(* Tests the contract between a caller's batch and a log exporter. *)
FUNCTION_BLOCK FB_TestLogExporters EXTENDS FB_TestSuite

THIS^.testExportSerializesWholeBatch();

(*
	export takes ownership of every record in the caller's batch and passes them to the serializer, so the
	caller holds nothing the exporter will release. Grouping by resource and scope is tested in FB_TestProtoJsonSerializer.
*)
METHOD testExportSerializesWholeBatch : REFERENCE TO FB_Test
VAR CONSTANT
	RECORD_COUNT: UDINT := 2;  // more than one, so the whole batch has to move, not just its head
END_VAR
VAR
	resource: FB_Resource(schemaUrl:='');
	provider: FB_LoggerProvider(resource:=resource);
	scope: FB_InstrumentationScope(name:='exporter.test', version:='1.0.0', schemaUrl:='');
	logger: FB_Logger(scope:=scope, provider:=provider);
	processor: FB_LogRecordProcessor_ForRecordsInspection(
		maxQueueSize:=0,
		scheduledDelayMillis:=1000,
		maxExportBatchSize:=512,
		exporter:=0
	);
	exporter: FB_LogRecordExporter_File_ForSerializationInspection;
	serialized: REFERENCE TO FB_LogRecordProtoJsonSerializer;
	emitSucceeded: BOOL;
	emitFailureReason: E_LoggerFailureReason;
	exporterFailureReason: E_LogRecordExporterFailureReason;
	exportSucceeded: BOOL;
	resourceLogs: SJsonValue;
	_idx: UDINT;
END_VAR
TcUnit.TEST('testExportSerializesWholeBatch');
	// arrange: the processor collects a batch emitted through the logger; its resource and scope do not matter here
	processor.free();
	FOR _idx := 1 TO RECORD_COUNT DO
		emitSucceeded := logger
			.startLogRecord(severityNumber:=E_SeverityNumber.INFO)
			.setTimestamp(TO_ULINT(_idx))
			.emit(failureResult=>emitFailureReason);
		THIS^.AssertTrue(emitSucceeded, 'Expected the logger to emit the record');
	END_FOR
	provider
		.stageProcessor(processor)
		.tick();
	THIS^.AssertEquals_UDINT(RECORD_COUNT, processor.records.count, 'Expected the processor to collect every emitted record');

	// act
	exportSucceeded := processor.exportRecords(exporter:=exporter, failureReason=>exporterFailureReason);

	// assert: the exporter owns the whole batch and serialized it
	THIS^.AssertTrue(
		exportSucceeded
		AND_THEN processor.records.count = 0
		AND_THEN exporterFailureReason = E_LogRecordExporterFailureReason.NA,
		'Expected export to succeed with no failure reason and take every record out of the batch'
	);
	serialized REF= exporter.serializer;
	resourceLogs := serialized.parser.FindMember(serialized.jsonValue, 'resourceLogs');
	THIS^.AssertTrue(resourceLogs <> 0 AND_THEN serialized.parser.IsArray(resourceLogs), 'Expected the exporter to serialize the batch into a resourceLogs array');

	exporter.free();
	processor.free();
TcUnit.TEST_FINISHED();
END_METHOD

END_FUNCTION_BLOCK

(* stored: Version 1.1.0.1
   POU FB_TestLogExporters: Id {6be9410b-9d69-4d16-a5fe-b31cbe727e6c}, SpecialFunc None
   Method testExportSerializesWholeBatch: Id {5d5f1575-5e45-48b1-b9ad-2eec80177025} *)
